Fanuc KAREL source: kb00176.KL

-- PROVISIONAL review KL for V1013-1; original PC SHA256 754970b2f864fce01f3975bbbd0ec889b0fe5ad6c4d51b779148ed52ad80e936
-- Incomplete behavior may be omitted. Consult companion uncertainty JSON. Do not deploy.
PROGRAM KB00176
%NOLOCKGROUP
BEGIN
  -- UNRESOLVED_PC offsets 5-12; opcodes 9D,23
  -- UNRESOLVED_PC offsets 17-32; opcodes 2E,22,32,35
  -- UNRESOLVED_PC offsets 37-44; opcodes 9D,23
  -- UNRESOLVED_PC offsets 49-79; opcodes 27,22,22,1C,22,27,9D,31
  -- UNRESOLVED_PC offsets 84-88; opcodes 7F
END KB00176
